(* Standard MKS 9XX series conversion *)
(* works for 925 *)
FUNCTION_BLOCK FB_9XX EXTENDS FB_GaugeBase
VAR_INPUT
END_VAR
VAR_OUTPUT
    {attribute 'pytmc' := '
    pv:
    '}
    PG	: ST_VG;
END_VAR
VAR_IN_OUT
END_VAR
VAR
    rV : REAL;
    fbGaugeState : FB_PressureState;
    rMaxPressure	:	REAL := 760; //Torr
    rMinPressure	:	REAL := 1E-5; //Torr
    rVMin : REAL:= 0.9;

    iTermBits: UINT := 30518 ; // The terminal's maximum value in bits default el3174 as per vacuum architecture
    (*IO*)
    i_iPRESS_R AT%I* :INT; // input Pressure // Link to analog Input
END_VAR

VAR CONSTANT
    (*Default set point 50 mT*)
    rDefaultVAC_SP: REAL := 5E-2;
END_VAR

(* Standard MKS 9XX series conversion *)
(* works for 972 and 925 *)


//Default setpoint
IF PG.rVAC_SP = 0 THEN
    PG.rVAC_SP := rDefaultVAC_SP;
END_IF
// check no div by zero
If (iTermBits=0) THEN iTermBits := 30518;END_IF
rV := 10*INT_TO_REAL(PG.i_iPRESS_R)/iTermBits;

IF rV >=rVMin THEN
    IF rV >= rVMin AND rV <= 1 THEN
        PG.rPRESS := 1E-5;
    ELSE
        PG.rPRESS := LREAL_TO_REAL(EXPT(10, rV-6));
    END_IF
    PG.xPRESS_OK := TRUE;
    PG.eState := Valid;
ELSE
    PG.xPRESS_OK := FALSE;
    IF (rV = 0) THEN PG.eState := GaugeDisconnected;
        ELSE  PG.eState := PressInvalid;
    END_IF
END_IF

(* Setpoint evaluation *)
PG.xAT_VAC := PG.xPRESS_OK AND (PG.rPRESS < PG.rVAC_SP);


(*Logger*)
ACT_Logger();
(*Soft IO Mapping*)
ACT_IO();

ACTION ACT_IO:
PG.i_iPRESS_R :=i_iPRESS_R;
PG.sPath := sPath;
END_ACTION

ACTION ACT_Logger:

//STATE Logger
IF ePrevState <> PG.eState THEN
      CASE PG.eState OF
        ValidHi:
            fbLogger(sMsg:='Gauge pressure valid high.', eSevr:=TcEventSeverity.Info);
        ValidLo:
            fbLogger(sMsg:='Gauge pressure valid low.', eSevr:=TcEventSeverity.Info);
        Valid:
            fbLogger(sMsg:='Gauge pressure valid.', eSevr:=TcEventSeverity.Info);
          GaugeDisconnected:
            fbLogger(sMsg:='Gauge Disconnected.', eSevr:=TcEventSeverity.Critical);
        PressInvalid:
            fbLogger(sMsg:='Gauge pressure invalid.', eSevr:=TcEventSeverity.Warning);
        OoR:
            fbLogger(sMsg:='Gauge pressure out of range.', eSevr:=TcEventSeverity.Warning);
        Starting:
            fbLogger(sMsg:='Gauge starting.', eSevr:=TcEventSeverity.Info);
      END_CASE
      ePrevState := PG.eState;
  END_IF
END_ACTION

METHOD M_SetBits : BOOL
VAR_INPUT
    TermBits : UINT; // The terminal's maximum value in bits
END_VAR
This^.iTermBits := TermBits;
END_METHOD

END_FUNCTION_BLOCK

(* stored: Version 1.1.0.1
   POU FB_9XX: Id {2b25be69-d890-49a3-9eed-41a1523a8d75}, SpecialFunc None
   Action ACT_IO: Id {fa0165d3-2f39-4dbf-b71c-224ecb928e0b}
   Action ACT_Logger: Id {8202116e-e944-4d2f-9609-fb14baf15925}
   Method M_SetBits: Id {c6390781-2f32-46e3-a37b-9fd31dd0725f} *)
